INTERFACE ITcoMessageProperties

METHOD Pin : ITcoMessageProperties
END_METHOD

PROPERTY Pinned : BOOL
GET
END_GET
END_PROPERTY

END_INTERFACE

(* stored: Version 1.1.0.1
   Itf ITcoMessageProperties: Id {033ac595-645d-056c-310a-5a8e070f1714}
   Method Pin: Id {54b58622-3387-07ec-2305-491e9eae5e49}
   Property Pinned: Id {dc7580a4-f337-0e34-06b3-f0bfdcc86bf6}
   Get Get: Id {787b8077-c24f-0b68-2628-9d2e00152a64} *)
